(****************************************************************************************************<br>
© Syntegon Group.<br>
All rights reserved, also regarding any disposal, exploitation, reproduction, editing, distribution,<br>
as well as in the event of applications for industrial property rights.<br>
*****************************************************************************************************<br>
DESCRIPTION:<br>
DEMO ONLY: independent sample applications side by side, for testing the gateway over ADS. All lines<br>
start at X = 0 and convey along +X. Each application is its own program:<br>
- P_VisuDemoDelta (Y = 0..1000): two infeeds, one outfeed, three Delta robots with different grippers; Infeed 1<br>
  is fed by a product generator and run, with Delta 1, by the sequence control P_VisuDemoMachine.<br>
- P_VisuDemoFxx (Y = 2500): an XTS loop above two belts evens out irregular gaps.<br>
- P_VisuDemoIdh (Y = 4100..4850): an XTS gantry picks in batches onto a tray belt.<br>
- P_VisuDemoCartesian (Y = 6500..7300): a Cartesian robot turns and tilts the products it places.<br>
- P_VisuDemoCartesianAxes (X = 4000, Y = 6500..7800): Cartesian robots without Y or without Z axis.<br>
- P_VisuDemoSpacing (Y = 9000): an XTS loop under one belt hands products back with a constant pitch.<br>
- P_VisuDemoStress (Y = 11000): load test with thousands of products, off unless DEMO_un_StressProducts is set.<br>
This program, called by PlcTask, sets the shared cycle time and fault phase (DEMO_GlobalVar), calls the machine's<br>
sequence control (recipe, commands, run state, machine messages: P_VisuDemoMachine) and then the applications.<br>
Part of the demo application Syn_Visu_Demo, which uses the Syn_Visu library like any machine project.<br>
****************************************************************************************************)
PROGRAM P_VisuDemo
VAR
	dn_TaskIndex						: DINT;
END_VAR

(****************************************************************************************************)
(* CYCLE TIME AND FAULT PHASE                                                                       *)
(****************************************************************************************************)
dn_TaskIndex := Tc2_System.GETCURTASKINDEXEX();
IF dn_TaskIndex > 0 THEN
	DEMO_GlobalVar.DEMO_lr_Dt := UDINT_TO_LREAL(TwinCAT_SystemInfoVarList._TaskInfo[dn_TaskIndex].CycleTime) * 1.0E-7;
ELSE
	DEMO_GlobalVar.DEMO_lr_Dt := 0.01;
END_IF
DEMO_GlobalVar.DEMO_lr_FaultPhase := DEMO_GlobalVar.DEMO_lr_FaultPhase + DEMO_GlobalVar.DEMO_lr_Dt;
IF DEMO_GlobalVar.DEMO_lr_FaultPhase >= DEMO_GlobalConst.DEMO_lr_FAULT_PERIOD THEN
	DEMO_GlobalVar.DEMO_lr_FaultPhase := DEMO_GlobalVar.DEMO_lr_FaultPhase - DEMO_GlobalConst.DEMO_lr_FAULT_PERIOD;
END_IF


(****************************************************************************************************)
(* MACHINE: recipe, commands and run state first, so the applications run with this cycle's values    *)
(****************************************************************************************************)
P_VisuDemoMachine();


(****************************************************************************************************)
(* APPLICATIONS                                                                                     *)
(****************************************************************************************************)
P_VisuDemoDelta();
P_VisuDemoFxx();
P_VisuDemoIdh();
P_VisuDemoCartesian();
P_VisuDemoCartesianAxes();
P_VisuDemoSpacing();
P_VisuDemoStress();

END_PROGRAM

(* stored: Version 1.1.0.1
   POU P_VisuDemo: Id {49b73753-a79a-401f-84bc-fc7827b66eb0}, SpecialFunc None *)
